(* IEC 61131-3 sources: ControlsBenchMUSE/codesys/library/examples/mappings/conveyor-m8, 8 files *)

(* ---- ST_CONV_Inputs.st ---- *)
TYPE ST_CONV_Inputs :
STRUCT
    // Generated by codesys/library/scripts/cb-map.mjs 0.1.0 from mappings/conveyor-m8.map.json; do not edit.
    // Raw inputs in native types; the session image carries them losslessly.
    PE_Entry : BOOL; // Digital[0]
    PE_D1Approach : BOOL; // Digital[1]
    PE_D2Approach : BOOL; // Digital[2]
    PE_ExitA : BOOL; // Digital[3]
    PE_ExitB : BOOL; // Digital[4]
    PE_Runout : BOOL; // Digital[5]
    D1_HomeFB : BOOL; // Digital[6]
    D1_ExtendedFB : BOOL; // Digital[7]
    D2_HomeFB : BOOL; // Digital[8]
    D2_ExtendedFB : BOOL; // Digital[9]
    Drive_RunningFB : BOOL; // Digital[10]
    Drive_Overload : BOOL; // Digital[11]
    ExitA_Ready : BOOL; // Digital[12]
    ExitB_Ready : BOOL; // Digital[13]
    Runout_Ready : BOOL; // Digital[14]
    Belt_SpeedActual : REAL; // Numeric.RealValue[0]
    Drive_Current : REAL; // Numeric.RealValue[1]
    D1_Position : REAL; // Numeric.RealValue[2]
    D2_Position : REAL; // Numeric.RealValue[3]
    Encoder_Count : UDINT; // Numeric.Unsigned[0], 32-bit
END_STRUCT
END_TYPE

(* ---- ST_CONV_Outputs.st ---- *)
TYPE ST_CONV_Outputs :
STRUCT
    // Generated by codesys/library/scripts/cb-map.mjs 0.1.0 from mappings/conveyor-m8.map.json; do not edit.
    // Application output commands in native types.
    Motor_RunCmd : BOOL; // Digital[0]
    D1_ExtendCmd : BOOL; // Digital[1]
    D2_ExtendCmd : BOOL; // Digital[2]
    StackLight_Red : BOOL; // Digital[3]
    StackLight_Green : BOOL; // Digital[4]
END_STRUCT
END_TYPE

(* ---- GVL_CONV_Map.st ---- *)
{attribute 'qualified_only'}
VAR_GLOBAL CONSTANT
    // Generated by codesys/library/scripts/cb-map.mjs 0.1.0 from mappings/conveyor-m8.map.json; do not edit.
    // Wire identities of this machine map.
    MAP_ID : STRING(32) := 'conveyor-m8';
    SCHEMA_ID : UDINT := 16#C69AC9A1; // raw input/output channel layout
    TAP_SCHEMA_ID : UDINT := 16#00000000; // observation tap list; 0 when none
    DEFAULT_DOMAIN_ID : UDINT := 1;
    TIMEOUT_US : ULINT := 500000;
END_VAR

(* ---- MAP_CONV_Config.st ---- *)
FUNCTION MAP_CONV_Config : CB.ST_CB_Config
VAR_INPUT
    DomainId : UDINT; // one value per authority domain in the application
END_VAR
VAR
    c : CB.ST_CB_Config;
END_VAR
// Generated by codesys/library/scripts/cb-map.mjs 0.1.0 from mappings/conveyor-m8.map.json; do not edit.
// Session configuration for this map.
c.DomainId := DomainId;
c.SchemaId := GVL_CONV_Map.SCHEMA_ID;
c.TimeoutUs := GVL_CONV_Map.TIMEOUT_US;
c.DigitalCount := 15;
c.SignedCount := 0;
c.UnsignedCount := 1;
c.RealCount := 4;
c.RealNonFiniteAllowed[0] := FALSE; // Belt_SpeedActual
c.RealNonFiniteAllowed[1] := FALSE; // Drive_Current
c.RealNonFiniteAllowed[2] := FALSE; // D1_Position
c.RealNonFiniteAllowed[3] := FALSE; // D2_Position
c.UnsignedBits[0] := 32; // Encoder_Count
MAP_CONV_Config := c;
END_FUNCTION

(* ---- MAP_CONV_PackInputs.st ---- *)
FUNCTION MAP_CONV_PackInputs : CB.ST_CB_Image
VAR_INPUT
    Source : ST_CONV_Inputs;
END_VAR
VAR
    image : CB.ST_CB_Image;
END_VAR
// Generated by codesys/library/scripts/cb-map.mjs 0.1.0 from mappings/conveyor-m8.map.json; do not edit.
// Raw acquisition into the session hardware image.
image.Digital[0] := Source.PE_Entry;
image.Digital[1] := Source.PE_D1Approach;
image.Digital[2] := Source.PE_D2Approach;
image.Digital[3] := Source.PE_ExitA;
image.Digital[4] := Source.PE_ExitB;
image.Digital[5] := Source.PE_Runout;
image.Digital[6] := Source.D1_HomeFB;
image.Digital[7] := Source.D1_ExtendedFB;
image.Digital[8] := Source.D2_HomeFB;
image.Digital[9] := Source.D2_ExtendedFB;
image.Digital[10] := Source.Drive_RunningFB;
image.Digital[11] := Source.Drive_Overload;
image.Digital[12] := Source.ExitA_Ready;
image.Digital[13] := Source.ExitB_Ready;
image.Digital[14] := Source.Runout_Ready;
image.Numeric.RealValue[0] := Source.Belt_SpeedActual;
image.Numeric.RealValue[1] := Source.Drive_Current;
image.Numeric.RealValue[2] := Source.D1_Position;
image.Numeric.RealValue[3] := Source.D2_Position;
image.Numeric.Unsigned[0] := Source.Encoder_Count;
MAP_CONV_PackInputs := image;
END_FUNCTION

(* ---- MAP_CONV_PackOutputs.st ---- *)
FUNCTION MAP_CONV_PackOutputs : CB.ST_CB_Image
VAR_INPUT
    Source : ST_CONV_Outputs;
END_VAR
VAR
    image : CB.ST_CB_Image;
END_VAR
// Generated by codesys/library/scripts/cb-map.mjs 0.1.0 from mappings/conveyor-m8.map.json; do not edit.
// Authentic commands into an output image for the DO/AO taps.
image.Digital[0] := Source.Motor_RunCmd;
image.Digital[1] := Source.D1_ExtendCmd;
image.Digital[2] := Source.D2_ExtendCmd;
image.Digital[3] := Source.StackLight_Red;
image.Digital[4] := Source.StackLight_Green;
MAP_CONV_PackOutputs := image;
END_FUNCTION

(* ---- MAP_CONV_UnpackInputs.st ---- *)
FUNCTION MAP_CONV_UnpackInputs : ST_CONV_Inputs
VAR_INPUT
    Image : CB.ST_CB_Image;
END_VAR
VAR
    values : ST_CONV_Inputs;
END_VAR
// Generated by codesys/library/scripts/cb-map.mjs 0.1.0 from mappings/conveyor-m8.map.json; do not edit.
// Selected image back to native types; the session has enforced each width.
values.PE_Entry := Image.Digital[0];
values.PE_D1Approach := Image.Digital[1];
values.PE_D2Approach := Image.Digital[2];
values.PE_ExitA := Image.Digital[3];
values.PE_ExitB := Image.Digital[4];
values.PE_Runout := Image.Digital[5];
values.D1_HomeFB := Image.Digital[6];
values.D1_ExtendedFB := Image.Digital[7];
values.D2_HomeFB := Image.Digital[8];
values.D2_ExtendedFB := Image.Digital[9];
values.Drive_RunningFB := Image.Digital[10];
values.Drive_Overload := Image.Digital[11];
values.ExitA_Ready := Image.Digital[12];
values.ExitB_Ready := Image.Digital[13];
values.Runout_Ready := Image.Digital[14];
values.Belt_SpeedActual := Image.Numeric.RealValue[0];
values.Drive_Current := Image.Numeric.RealValue[1];
values.D1_Position := Image.Numeric.RealValue[2];
values.D2_Position := Image.Numeric.RealValue[3];
values.Encoder_Count := Image.Numeric.Unsigned[0];
MAP_CONV_UnpackInputs := values;
END_FUNCTION

(* ---- MAP_CONV_UnpackOutputs.st ---- *)
FUNCTION MAP_CONV_UnpackOutputs : ST_CONV_Outputs
VAR_INPUT
    Image : CB.ST_CB_Image;
END_VAR
VAR
    values : ST_CONV_Outputs;
END_VAR
// Generated by codesys/library/scripts/cb-map.mjs 0.1.0 from mappings/conveyor-m8.map.json; do not edit.
// Physical sink values; configured SuppressedValues must fit each native type.
values.Motor_RunCmd := Image.Digital[0];
values.D1_ExtendCmd := Image.Digital[1];
values.D2_ExtendCmd := Image.Digital[2];
values.StackLight_Red := Image.Digital[3];
values.StackLight_Green := Image.Digital[4];
MAP_CONV_UnpackOutputs := values;
END_FUNCTION
